(* IEC 61131-3 sources: trust-platform/examples/OSCAT/tank_farm_transfer_skid/oop/src, 3 files *)

(* ---- Main.st ---- *)
(* Pattern role: IPlantNode is the contract boundary for the Composite and Iterator example. *)
INTERFACE IPlantNode EXTENDS IComponent
    PROPERTY NodeId : INT
    GET
    END_GET
    END_PROPERTY

    PROPERTY ChildCount : INT
    GET
    END_GET
    END_PROPERTY

    PROPERTY StoppedCount : INT
    GET
    END_GET
    END_PROPERTY

    PROPERTY AlarmCount : INT
    GET
    END_GET
    END_PROPERTY

    METHOD GetChild : IPlantNode
    VAR_INPUT
        Index : INT;
    END_VAR
    END_METHOD

    METHOD EmergencyStop
    END_METHOD

    METHOD AcknowledgeAll
    END_METHOD
END_INTERFACE

(* Pattern role: TankNode is a concrete implementation in the Composite and Iterator example. *)
FUNCTION_BLOCK TankNode IMPLEMENTS IPlantNode
VAR
    NodeIdValue : INT;
    StoppedValue : BOOL;
    AlarmValue : BOOL;
    AckCountValue : INT;
    ReadyValue : BOOL;
    ErrorValue : BOOL;
    ErrorIdValue : WORD;
    StatusValue : BYTE;
    LevelFilter : Pt1Filter;
    HighAlarm : HysteresisSwitch;
    AlarmLimits : RealRange;
END_VAR

METHOD PUBLIC Configure
VAR_INPUT
    NodeId : INT;
    HighAlarmActive : BOOL;
END_VAR
NodeIdValue := NodeId;
AlarmValue := HighAlarmActive;
END_METHOD

METHOD PUBLIC Initialize
ReadyValue := TRUE;
LevelFilter.Initialize();
LevelFilter.Configure(TimeConstant := T#1s, Gain := REAL#1.0);
AlarmLimits.Low := REAL#5.0;
AlarmLimits.High := REAL#90.0;
HighAlarm.Initialize();
HighAlarm.SetLimits(Limits := AlarmLimits);
ClearError();
END_METHOD

METHOD PUBLIC Reset
StoppedValue := FALSE;
AckCountValue := INT#0;
ClearError();
END_METHOD

METHOD PUBLIC ClearError
ErrorValue := FALSE;
ErrorIdValue := WORD#0;
StatusValue := BYTE#0;
END_METHOD

METHOD PUBLIC Snapshot : ComponentStatus
VAR
    Result : ComponentStatus;
END_VAR
Result.Ready := ReadyValue;
Result.Error := ErrorValue;
Result.ErrorId := ErrorIdValue;
Result.Status := StatusValue;
Snapshot := Result;
END_METHOD

METHOD PUBLIC UpdateLevel
VAR_INPUT
    LevelPct : REAL;
END_VAR
AlarmValue := HighAlarm.Update(MeasuredValue := LevelFilter.Update(Sample := LevelPct));
END_METHOD

METHOD PUBLIC GetChild : IPlantNode
VAR_INPUT
    Index : INT;
END_VAR
GetChild := THIS;
END_METHOD

METHOD PUBLIC EmergencyStop
StoppedValue := TRUE;
END_METHOD

METHOD PUBLIC AcknowledgeAll
IF AlarmValue THEN
    AckCountValue := AckCountValue + INT#1;
END_IF;
AlarmValue := FALSE;
END_METHOD

PUBLIC PROPERTY NodeId : INT
GET
    NodeId := NodeIdValue;
END_GET
END_PROPERTY

PUBLIC PROPERTY ChildCount : INT
GET
    ChildCount := INT#0;
END_GET
END_PROPERTY

PUBLIC PROPERTY StoppedCount : INT
GET
    IF StoppedValue THEN
        StoppedCount := INT#1;
    ELSE
        StoppedCount := INT#0;
    END_IF;
END_GET
END_PROPERTY

PUBLIC PROPERTY AlarmCount : INT
GET
    IF AlarmValue THEN
        AlarmCount := INT#1;
    ELSE
        AlarmCount := INT#0;
    END_IF;
END_GET
END_PROPERTY

PUBLIC PROPERTY Ready : BOOL
GET
    Ready := ReadyValue;
END_GET
END_PROPERTY

PUBLIC PROPERTY Error : BOOL
GET
    Error := ErrorValue;
END_GET
END_PROPERTY

PUBLIC PROPERTY ErrorId : WORD
GET
    ErrorId := ErrorIdValue;
END_GET
END_PROPERTY

PUBLIC PROPERTY Status : BYTE
GET
    Status := StatusValue;
END_GET
END_PROPERTY
END_FUNCTION_BLOCK

(* Pattern role: AreaNode is a concrete implementation in the Composite and Iterator example. *)
FUNCTION_BLOCK AreaNode IMPLEMENTS IPlantNode
VAR
    NodeIdValue : INT;
    Tank1 : TankNode;
    Tank2 : TankNode;
    ReadyValue : BOOL;
    ErrorValue : BOOL;
    ErrorIdValue : WORD;
    StatusValue : BYTE;
END_VAR

METHOD PUBLIC Configure
VAR_INPUT
    NodeId : INT;
    Tank1Alarm : BOOL;
    Tank2Alarm : BOOL;
END_VAR
NodeIdValue := NodeId;
Tank1.Configure(NodeId := NodeId * INT#10 + INT#1, HighAlarmActive := Tank1Alarm);
Tank2.Configure(NodeId := NodeId * INT#10 + INT#2, HighAlarmActive := Tank2Alarm);
END_METHOD

METHOD PUBLIC Initialize
ReadyValue := TRUE;
Tank1.Initialize();
Tank2.Initialize();
ClearError();
END_METHOD

METHOD PUBLIC Reset
Tank1.Reset();
Tank2.Reset();
ClearError();
END_METHOD

METHOD PUBLIC ClearError
ErrorValue := FALSE;
ErrorIdValue := WORD#0;
StatusValue := BYTE#0;
END_METHOD

METHOD PUBLIC Snapshot : ComponentStatus
VAR
    Result : ComponentStatus;
END_VAR
Result.Ready := ReadyValue;
Result.Error := ErrorValue;
Result.ErrorId := ErrorIdValue;
Result.Status := StatusValue;
Snapshot := Result;
END_METHOD

METHOD PUBLIC GetChild : IPlantNode
VAR_INPUT
    Index : INT;
END_VAR
IF Index = INT#1 THEN
    GetChild := Tank1;
ELSE
    GetChild := Tank2;
END_IF;
END_METHOD

METHOD PUBLIC EmergencyStop
Tank1.EmergencyStop();
Tank2.EmergencyStop();
END_METHOD

METHOD PUBLIC AcknowledgeAll
Tank1.AcknowledgeAll();
Tank2.AcknowledgeAll();
END_METHOD

PUBLIC PROPERTY NodeId : INT
GET
    NodeId := NodeIdValue;
END_GET
END_PROPERTY

PUBLIC PROPERTY ChildCount : INT
GET
    ChildCount := INT#2;
END_GET
END_PROPERTY

PUBLIC PROPERTY StoppedCount : INT
GET
    StoppedCount := Tank1.StoppedCount + Tank2.StoppedCount;
END_GET
END_PROPERTY

PUBLIC PROPERTY AlarmCount : INT
GET
    AlarmCount := Tank1.AlarmCount + Tank2.AlarmCount;
END_GET
END_PROPERTY

PUBLIC PROPERTY Ready : BOOL
GET
    Ready := ReadyValue;
END_GET
END_PROPERTY

PUBLIC PROPERTY Error : BOOL
GET
    Error := ErrorValue;
END_GET
END_PROPERTY

PUBLIC PROPERTY ErrorId : WORD
GET
    ErrorId := ErrorIdValue;
END_GET
END_PROPERTY

PUBLIC PROPERTY Status : BYTE
GET
    Status := StatusValue;
END_GET
END_PROPERTY
END_FUNCTION_BLOCK

(* Pattern role: FarmNode is a concrete implementation in the Composite and Iterator example. *)
FUNCTION_BLOCK FarmNode IMPLEMENTS IPlantNode
VAR
    Area1 : AreaNode;
    Area2 : AreaNode;
    ReadyValue : BOOL;
    ErrorValue : BOOL;
    ErrorIdValue : WORD;
    StatusValue : BYTE;
END_VAR

METHOD PUBLIC Initialize
ReadyValue := TRUE;
Area1.Initialize();
Area2.Initialize();
Area1.Configure(NodeId := INT#1, Tank1Alarm := TRUE, Tank2Alarm := FALSE);
Area2.Configure(NodeId := INT#2, Tank1Alarm := FALSE, Tank2Alarm := TRUE);
ClearError();
END_METHOD

METHOD PUBLIC Reset
Area1.Reset();
Area2.Reset();
ClearError();
END_METHOD

METHOD PUBLIC ClearError
ErrorValue := FALSE;
ErrorIdValue := WORD#0;
StatusValue := BYTE#0;
END_METHOD

METHOD PUBLIC Snapshot : ComponentStatus
VAR
    Result : ComponentStatus;
END_VAR
Result.Ready := ReadyValue;
Result.Error := ErrorValue;
Result.ErrorId := ErrorIdValue;
Result.Status := StatusValue;
Snapshot := Result;
END_METHOD

METHOD PUBLIC GetChild : IPlantNode
VAR_INPUT
    Index : INT;
END_VAR
IF Index = INT#1 THEN
    GetChild := Area1;
ELSE
    GetChild := Area2;
END_IF;
END_METHOD

METHOD PUBLIC EmergencyStop
Area1.EmergencyStop();
Area2.EmergencyStop();
END_METHOD

METHOD PUBLIC AcknowledgeAll
Area1.AcknowledgeAll();
Area2.AcknowledgeAll();
END_METHOD

METHOD PUBLIC EmergencyStopArea
VAR_INPUT
    AreaIndex : INT;
END_VAR
VAR
    Area : IPlantNode;
END_VAR
Area := GetChild(Index := AreaIndex);
Area.EmergencyStop();
END_METHOD

PUBLIC PROPERTY NodeId : INT
GET
    NodeId := INT#100;
END_GET
END_PROPERTY

PUBLIC PROPERTY ChildCount : INT
GET
    ChildCount := INT#2;
END_GET
END_PROPERTY

PUBLIC PROPERTY StoppedCount : INT
GET
    StoppedCount := Area1.StoppedCount + Area2.StoppedCount;
END_GET
END_PROPERTY

PUBLIC PROPERTY AlarmCount : INT
GET
    AlarmCount := Area1.AlarmCount + Area2.AlarmCount;
END_GET
END_PROPERTY

PUBLIC PROPERTY Ready : BOOL
GET
    Ready := ReadyValue;
END_GET
END_PROPERTY

PUBLIC PROPERTY Error : BOOL
GET
    Error := ErrorValue;
END_GET
END_PROPERTY

PUBLIC PROPERTY ErrorId : WORD
GET
    ErrorId := ErrorIdValue;
END_GET
END_PROPERTY

PUBLIC PROPERTY Status : BYTE
GET
    Status := StatusValue;
END_GET
END_PROPERTY
END_FUNCTION_BLOCK

(* Scan role: Main wires the example objects and exposes the PLC call path under test. *)
PROGRAM Main
VAR
    Farm : FarmNode;
    Area : IPlantNode;
    Tank : IPlantNode;
    AreaStopCommand : BOOL;
    AreaIndex : INT;
    TankIndex : INT;
    TotalTankAlarms : INT;
    AreaStoppedOut : BOOL;
END_VAR

Farm.Initialize();
IF AreaStopCommand THEN
    Farm.EmergencyStopArea(AreaIndex := AreaIndex);
END_IF;
TotalTankAlarms := INT#0;
FOR AreaIndex := INT#1 TO Farm.ChildCount DO
    Area := Farm.GetChild(Index := AreaIndex);
    FOR TankIndex := INT#1 TO Area.ChildCount DO
        Tank := Area.GetChild(Index := TankIndex);
        TotalTankAlarms := TotalTankAlarms + Tank.AlarmCount;
    END_FOR;
END_FOR;
AreaStoppedOut := Farm.StoppedCount > INT#0;
END_PROGRAM

(* ---- Configuration.st ---- *)
CONFIGURATION TankFarmOopConfiguration
RESOURCE TankFarmOop ON PLC
    TASK MainTask (INTERVAL := T#100ms, PRIORITY := 1);
    PROGRAM Farm WITH MainTask : Main;
END_RESOURCE
VAR_CONFIG
    Farm.AreaStopCommand AT %IX0.0 : BOOL;
    Farm.AreaIndex AT %IW2 : INT;
    Farm.AreaStoppedOut AT %QX0.0 : BOOL;
END_VAR
END_CONFIGURATION

(* ---- Tests.st ---- *)
TEST_PROGRAM TankFarmCompositeStopsOneAreaThroughPlantNode
VAR
    Farm : FarmNode;
    Area : IPlantNode;
    Tank : IPlantNode;
END_VAR

Farm.Initialize();
ASSERT_EQUAL(EXPECTED := INT#2, ACTUAL := Farm.ChildCount);
Area := Farm.GetChild(Index := INT#2);
ASSERT_EQUAL(EXPECTED := INT#2, ACTUAL := Area.ChildCount);
Tank := Area.GetChild(Index := INT#1);
ASSERT_EQUAL(EXPECTED := INT#0, ACTUAL := Farm.StoppedCount);

Area.EmergencyStop();
ASSERT_EQUAL(EXPECTED := INT#2, ACTUAL := Farm.StoppedCount);
ASSERT_EQUAL(EXPECTED := INT#1, ACTUAL := Tank.StoppedCount);
END_TEST_PROGRAM

TEST_PROGRAM TankFarmCompositeAcknowledgesAlarmTree
VAR
    Farm : FarmNode;
END_VAR

Farm.Initialize();
ASSERT_EQUAL(EXPECTED := INT#2, ACTUAL := Farm.AlarmCount);
Farm.AcknowledgeAll();
ASSERT_EQUAL(EXPECTED := INT#0, ACTUAL := Farm.AlarmCount);
END_TEST_PROGRAM

(* Per-area isolation test: drives EmergencyStop on one area only and
   verifies that the OTHER area's tanks remain unaffected. Catches
   bugs where the composite's recursion descends into the wrong subtree
   or where StoppedCount accumulates beyond the affected subtree. *)
TEST_PROGRAM TankFarmEmergencyStopIsLocalToOneAreaOnly
VAR
    Farm : FarmNode;
    Area1 : IPlantNode;
    Area2 : IPlantNode;
    Tank1Of2 : IPlantNode;
END_VAR

Farm.Initialize();

(* Stop Area 2 only - Area 2's tanks count as stopped *)
Area2 := Farm.GetChild(Index := INT#2);
Area2.EmergencyStop();
ASSERT_EQUAL(EXPECTED := INT#2, ACTUAL := Farm.StoppedCount);

(* Area 1 must NOT be stopped - the recursion stays within the called
   subtree and does not cross into siblings *)
Area1 := Farm.GetChild(Index := INT#1);
Tank1Of2 := Area2.GetChild(Index := INT#1);
ASSERT_EQUAL(EXPECTED := INT#1, ACTUAL := Tank1Of2.StoppedCount);
END_TEST_PROGRAM

(* Iterator boundary: traversal across all areas and tanks in the farm
   matches the manual aggregation. Catches regressions where ChildCount
   reports the wrong count or GetChild returns the wrong node. *)
TEST_PROGRAM TankFarmIteratorVisitsEveryLeafExactlyOnce
VAR
    Farm : FarmNode;
    Area : IPlantNode;
    Tank : IPlantNode;
    AreaIndex : INT;
    TankIndex : INT;
    LeafCount : INT;
    AlarmTotal : INT;
END_VAR

Farm.Initialize();
LeafCount := INT#0;
AlarmTotal := INT#0;
FOR AreaIndex := INT#1 TO Farm.ChildCount DO
    Area := Farm.GetChild(Index := AreaIndex);
    FOR TankIndex := INT#1 TO Area.ChildCount DO
        Tank := Area.GetChild(Index := TankIndex);
        LeafCount := LeafCount + INT#1;
        AlarmTotal := AlarmTotal + Tank.AlarmCount;
    END_FOR;
END_FOR;
(* 2 areas x 2 tanks = 4 leaves *)
ASSERT_EQUAL(EXPECTED := INT#4, ACTUAL := LeafCount);
(* Aggregated leaf alarms must equal the farm's aggregated alarm count *)
ASSERT_EQUAL(EXPECTED := AlarmTotal, ACTUAL := Farm.AlarmCount);
END_TEST_PROGRAM

(* Per-leaf isolation: acknowledging a single tank's alarm must not
   touch the alarm state of other tanks in the same area or in other
   areas. *)
TEST_PROGRAM TankFarmPerLeafAcknowledgeIsLocal
VAR
    Farm : FarmNode;
    Area1 : IPlantNode;
    Tank1Of1 : IPlantNode;
END_VAR

Farm.Initialize();
(* Initial setup: Area1.Tank1 has alarm; Area2.Tank2 has alarm; total = 2 *)
ASSERT_EQUAL(EXPECTED := INT#2, ACTUAL := Farm.AlarmCount);

(* Acknowledge only Area1.Tank1 - the alarm in Area2.Tank2 must remain *)
Area1 := Farm.GetChild(Index := INT#1);
Tank1Of1 := Area1.GetChild(Index := INT#1);
Tank1Of1.AcknowledgeAll();
(* Total drops to 1 - the other alarm is still pending *)
ASSERT_EQUAL(EXPECTED := INT#1, ACTUAL := Farm.AlarmCount);
END_TEST_PROGRAM

(* Recursive EmergencyStop on the root farm node stops every leaf. *)
TEST_PROGRAM TankFarmRootEmergencyStopStopsAllLeaves
VAR
    Farm : FarmNode;
END_VAR

Farm.Initialize();
ASSERT_EQUAL(EXPECTED := INT#0, ACTUAL := Farm.StoppedCount);

Farm.EmergencyStop();
(* All four leaves must now report stopped *)
ASSERT_EQUAL(EXPECTED := INT#4, ACTUAL := Farm.StoppedCount);
END_TEST_PROGRAM

(* Per-FB isolation: two FarmNode instances must keep independent
   stop/alarm state. Catches a class of bug where shared state leaks
   between composite instances. *)
TEST_PROGRAM TankFarmFarmNodeInstancesAreIndependent
VAR
    FarmA : FarmNode;
    FarmB : FarmNode;
END_VAR

FarmA.Initialize();
FarmB.Initialize();

(* Stop FarmA only; FarmB unchanged *)
FarmA.EmergencyStop();
ASSERT_EQUAL(EXPECTED := INT#4, ACTUAL := FarmA.StoppedCount);
ASSERT_EQUAL(EXPECTED := INT#0, ACTUAL := FarmB.StoppedCount);

(* Acknowledge FarmB; FarmA's alarms unchanged *)
FarmB.AcknowledgeAll();
ASSERT_EQUAL(EXPECTED := INT#0, ACTUAL := FarmB.AlarmCount);
ASSERT_EQUAL(EXPECTED := INT#2, ACTUAL := FarmA.AlarmCount);
END_TEST_PROGRAM

(* EmergencyStopArea using the typed helper produces the same effect as
   walking the tree manually with GetChild + EmergencyStop. *)
TEST_PROGRAM TankFarmEmergencyStopAreaMatchesManualWalk
VAR
    Farm : FarmNode;
    AreaA : IPlantNode;
END_VAR

Farm.Initialize();
Farm.EmergencyStopArea(AreaIndex := INT#1);
(* Both tanks in Area 1 are stopped *)
AreaA := Farm.GetChild(Index := INT#1);
ASSERT_EQUAL(EXPECTED := INT#2, ACTUAL := AreaA.StoppedCount);
(* Area 2 untouched *)
ASSERT_EQUAL(EXPECTED := INT#2, ACTUAL := Farm.StoppedCount);
END_TEST_PROGRAM
